TYPE "st_Io_Ph_DigitalOutputs"
VERSION : 0.1
   STRUCT
      Zone1_K7k5Ss_Close { ExternalAccessible := 'False'; ExternalVisible := 'False'; ExternalWritable := 'False'; S7_SetPoint := 'False'} : "st_Io_Ph_DigitalOutput";
      Zone1_K7k5Vfd_Close { ExternalAccessible := 'False'; ExternalVisible := 'False'; ExternalWritable := 'False'; S7_SetPoint := 'False'} : "st_Io_Ph_DigitalOutput";
      Zone1_K37Ss_Close { ExternalAccessible := 'False'; ExternalVisible := 'False'; ExternalWritable := 'False'; S7_SetPoint := 'False'} : "st_Io_Ph_DigitalOutput";
      Zone1_K37Vfd_Close { ExternalAccessible := 'False'; ExternalVisible := 'False'; ExternalWritable := 'False'; S7_SetPoint := 'False'} : "st_Io_Ph_DigitalOutput";
      Zone1_K110Ss_Close { ExternalAccessible := 'False'; ExternalVisible := 'False'; ExternalWritable := 'False'; S7_SetPoint := 'False'} : "st_Io_Ph_DigitalOutput";
      Zone1_K110Vfd_Close { ExternalAccessible := 'False'; ExternalVisible := 'False'; ExternalWritable := 'False'; S7_SetPoint := 'False'} : "st_Io_Ph_DigitalOutput";
      Zone1_Q560Ss_Open { ExternalAccessible := 'False'; ExternalVisible := 'False'; ExternalWritable := 'False'; S7_SetPoint := 'False'} : "st_Io_Ph_DigitalOutput";
      Zone1_Q560Ss_Close { ExternalAccessible := 'False'; ExternalVisible := 'False'; ExternalWritable := 'False'; S7_SetPoint := 'False'} : "st_Io_Ph_DigitalOutput";
      Zone1_Q560Ss_ChargeSpring { ExternalAccessible := 'False'; ExternalVisible := 'False'; ExternalWritable := 'False'; S7_SetPoint := 'False'} : "st_Io_Ph_DigitalOutput";
      Zone1_Q630Vfd_Open { ExternalAccessible := 'False'; ExternalVisible := 'False'; ExternalWritable := 'False'; S7_SetPoint := 'False'} : "st_Io_Ph_DigitalOutput";
      Zone1_Q630Vfd_Close { ExternalAccessible := 'False'; ExternalVisible := 'False'; ExternalWritable := 'False'; S7_SetPoint := 'False'} : "st_Io_Ph_DigitalOutput";
      Zone1_Q630Vfd_ChargeSpring { ExternalAccessible := 'False'; ExternalVisible := 'False'; ExternalWritable := 'False'; S7_SetPoint := 'False'} : "st_Io_Ph_DigitalOutput";
      Zone1_LampGreen { ExternalAccessible := 'False'; ExternalVisible := 'False'; ExternalWritable := 'False'; S7_SetPoint := 'False'} : "st_Io_Ph_DigitalOutput";
      Zone1_LampYellow { ExternalAccessible := 'False'; ExternalVisible := 'False'; ExternalWritable := 'False'; S7_SetPoint := 'False'} : "st_Io_Ph_DigitalOutput";
      Zone1_LampRed { ExternalAccessible := 'False'; ExternalVisible := 'False'; ExternalWritable := 'False'; S7_SetPoint := 'False'} : "st_Io_Ph_DigitalOutput";
      Zone1_LampStart { ExternalAccessible := 'False'; ExternalVisible := 'False'; ExternalWritable := 'False'; S7_SetPoint := 'False'} : "st_Io_Ph_DigitalOutput";
      Zone1_LampStop { ExternalAccessible := 'False'; ExternalVisible := 'False'; ExternalWritable := 'False'; S7_SetPoint := 'False'} : "st_Io_Ph_DigitalOutput";
      Zone1_LampTakeSample { ExternalAccessible := 'False'; ExternalVisible := 'False'; ExternalWritable := 'False'; S7_SetPoint := 'False'} : "st_Io_Ph_DigitalOutput";
      Zone1_LampEStop { ExternalAccessible := 'False'; ExternalVisible := 'False'; ExternalWritable := 'False'; S7_SetPoint := 'False'} : "st_Io_Ph_DigitalOutput";
      Zone1_LampPanelEStop { ExternalAccessible := 'False'; ExternalVisible := 'False'; ExternalWritable := 'False'; S7_SetPoint := 'False'} : "st_Io_Ph_DigitalOutput";
      Zone2_K7k5Ss_Close { ExternalAccessible := 'False'; ExternalVisible := 'False'; ExternalWritable := 'False'; S7_SetPoint := 'False'} : "st_Io_Ph_DigitalOutput";
      Zone2_K7k5Vfd_Close { ExternalAccessible := 'False'; ExternalVisible := 'False'; ExternalWritable := 'False'; S7_SetPoint := 'False'} : "st_Io_Ph_DigitalOutput";
      Zone2_K37Ss_Close { ExternalAccessible := 'False'; ExternalVisible := 'False'; ExternalWritable := 'False'; S7_SetPoint := 'False'} : "st_Io_Ph_DigitalOutput";
      Zone2_K37Vfd_Close { ExternalAccessible := 'False'; ExternalVisible := 'False'; ExternalWritable := 'False'; S7_SetPoint := 'False'} : "st_Io_Ph_DigitalOutput";
      Zone2_K110Ss_Close { ExternalAccessible := 'False'; ExternalVisible := 'False'; ExternalWritable := 'False'; S7_SetPoint := 'False'} : "st_Io_Ph_DigitalOutput";
      Zone2_K110Vfd_Close { ExternalAccessible := 'False'; ExternalVisible := 'False'; ExternalWritable := 'False'; S7_SetPoint := 'False'} : "st_Io_Ph_DigitalOutput";
      Zone2_Q560Ss_Open { ExternalAccessible := 'False'; ExternalVisible := 'False'; ExternalWritable := 'False'; S7_SetPoint := 'False'} : "st_Io_Ph_DigitalOutput";
      Zone2_Q560Ss_Close { ExternalAccessible := 'False'; ExternalVisible := 'False'; ExternalWritable := 'False'; S7_SetPoint := 'False'} : "st_Io_Ph_DigitalOutput";
      Zone2_Q560Ss_ChargeSpring { ExternalAccessible := 'False'; ExternalVisible := 'False'; ExternalWritable := 'False'; S7_SetPoint := 'False'} : "st_Io_Ph_DigitalOutput";
      Zone2_Q630Vfd_Open { ExternalAccessible := 'False'; ExternalVisible := 'False'; ExternalWritable := 'False'; S7_SetPoint := 'False'} : "st_Io_Ph_DigitalOutput";
      Zone2_Q630Vfd_Close { ExternalAccessible := 'False'; ExternalVisible := 'False'; ExternalWritable := 'False'; S7_SetPoint := 'False'} : "st_Io_Ph_DigitalOutput";
      Zone2_Q630Vfd_ChargeSpring { ExternalAccessible := 'False'; ExternalVisible := 'False'; ExternalWritable := 'False'; S7_SetPoint := 'False'} : "st_Io_Ph_DigitalOutput";
      Zone2_LampGreen { ExternalAccessible := 'False'; ExternalVisible := 'False'; ExternalWritable := 'False'; S7_SetPoint := 'False'} : "st_Io_Ph_DigitalOutput";
      Zone2_LampYellow { ExternalAccessible := 'False'; ExternalVisible := 'False'; ExternalWritable := 'False'; S7_SetPoint := 'False'} : "st_Io_Ph_DigitalOutput";
      Zone2_LampRed { ExternalAccessible := 'False'; ExternalVisible := 'False'; ExternalWritable := 'False'; S7_SetPoint := 'False'} : "st_Io_Ph_DigitalOutput";
      Zone2_LampStart { ExternalAccessible := 'False'; ExternalVisible := 'False'; ExternalWritable := 'False'; S7_SetPoint := 'False'} : "st_Io_Ph_DigitalOutput";
      Zone2_LampStop { ExternalAccessible := 'False'; ExternalVisible := 'False'; ExternalWritable := 'False'; S7_SetPoint := 'False'} : "st_Io_Ph_DigitalOutput";
      Zone2_LampTakeSample { ExternalAccessible := 'False'; ExternalVisible := 'False'; ExternalWritable := 'False'; S7_SetPoint := 'False'} : "st_Io_Ph_DigitalOutput";
      Zone2_LampEStop { ExternalAccessible := 'False'; ExternalVisible := 'False'; ExternalWritable := 'False'; S7_SetPoint := 'False'} : "st_Io_Ph_DigitalOutput";
      Zone2_LampPanelEStop { ExternalAccessible := 'False'; ExternalVisible := 'False'; ExternalWritable := 'False'; S7_SetPoint := 'False'} : "st_Io_Ph_DigitalOutput";
      Zone3_K7k5Ss_Close { ExternalAccessible := 'False'; ExternalVisible := 'False'; ExternalWritable := 'False'; S7_SetPoint := 'False'} : "st_Io_Ph_DigitalOutput";
      Zone3_K7k5Vfd_Close { ExternalAccessible := 'False'; ExternalVisible := 'False'; ExternalWritable := 'False'; S7_SetPoint := 'False'} : "st_Io_Ph_DigitalOutput";
      Zone3_K37Ss_Close { ExternalAccessible := 'False'; ExternalVisible := 'False'; ExternalWritable := 'False'; S7_SetPoint := 'False'} : "st_Io_Ph_DigitalOutput";
      Zone3_K37Vfd_Close { ExternalAccessible := 'False'; ExternalVisible := 'False'; ExternalWritable := 'False'; S7_SetPoint := 'False'} : "st_Io_Ph_DigitalOutput";
      Zone3_K110Ss_Close { ExternalAccessible := 'False'; ExternalVisible := 'False'; ExternalWritable := 'False'; S7_SetPoint := 'False'} : "st_Io_Ph_DigitalOutput";
      Zone3_K110Vfd_Close { ExternalAccessible := 'False'; ExternalVisible := 'False'; ExternalWritable := 'False'; S7_SetPoint := 'False'} : "st_Io_Ph_DigitalOutput";
      Zone3_Q560Ss_Open { ExternalAccessible := 'False'; ExternalVisible := 'False'; ExternalWritable := 'False'; S7_SetPoint := 'False'} : "st_Io_Ph_DigitalOutput";
      Zone3_Q560Ss_Close { ExternalAccessible := 'False'; ExternalVisible := 'False'; ExternalWritable := 'False'; S7_SetPoint := 'False'} : "st_Io_Ph_DigitalOutput";
      Zone3_Q560Ss_ChargeSpring { ExternalAccessible := 'False'; ExternalVisible := 'False'; ExternalWritable := 'False'; S7_SetPoint := 'False'} : "st_Io_Ph_DigitalOutput";
      Zone3_Q630Vfd_Open { ExternalAccessible := 'False'; ExternalVisible := 'False'; ExternalWritable := 'False'; S7_SetPoint := 'False'} : "st_Io_Ph_DigitalOutput";
      Zone3_Q630Vfd_Close { ExternalAccessible := 'False'; ExternalVisible := 'False'; ExternalWritable := 'False'; S7_SetPoint := 'False'} : "st_Io_Ph_DigitalOutput";
      Zone3_Q630Vfd_ChargeSpring { ExternalAccessible := 'False'; ExternalVisible := 'False'; ExternalWritable := 'False'; S7_SetPoint := 'False'} : "st_Io_Ph_DigitalOutput";
      Zone3_LampGreen { ExternalAccessible := 'False'; ExternalVisible := 'False'; ExternalWritable := 'False'; S7_SetPoint := 'False'} : "st_Io_Ph_DigitalOutput";
      Zone3_LampYellow { ExternalAccessible := 'False'; ExternalVisible := 'False'; ExternalWritable := 'False'; S7_SetPoint := 'False'} : "st_Io_Ph_DigitalOutput";
      Zone3_LampRed { ExternalAccessible := 'False'; ExternalVisible := 'False'; ExternalWritable := 'False'; S7_SetPoint := 'False'} : "st_Io_Ph_DigitalOutput";
      Zone3_LampStart { ExternalAccessible := 'False'; ExternalVisible := 'False'; ExternalWritable := 'False'; S7_SetPoint := 'False'} : "st_Io_Ph_DigitalOutput";
      Zone3_LampStop { ExternalAccessible := 'False'; ExternalVisible := 'False'; ExternalWritable := 'False'; S7_SetPoint := 'False'} : "st_Io_Ph_DigitalOutput";
      Zone3_LampTakeSample { ExternalAccessible := 'False'; ExternalVisible := 'False'; ExternalWritable := 'False'; S7_SetPoint := 'False'} : "st_Io_Ph_DigitalOutput";
      Zone3_LampEStop { ExternalAccessible := 'False'; ExternalVisible := 'False'; ExternalWritable := 'False'; S7_SetPoint := 'False'} : "st_Io_Ph_DigitalOutput";
      Zone3_LampPanelEStop { ExternalAccessible := 'False'; ExternalVisible := 'False'; ExternalWritable := 'False'; S7_SetPoint := 'False'} : "st_Io_Ph_DigitalOutput";
      Drive_7k5Ss_Run { ExternalAccessible := 'False'; ExternalVisible := 'False'; ExternalWritable := 'False'; S7_SetPoint := 'False'} : "st_Io_Ph_DigitalOutput";
      Drive_7k5Vfd_Run { ExternalAccessible := 'False'; ExternalVisible := 'False'; ExternalWritable := 'False'; S7_SetPoint := 'False'} : "st_Io_Ph_DigitalOutput";
      Drive_37Ss_Run { ExternalAccessible := 'False'; ExternalVisible := 'False'; ExternalWritable := 'False'; S7_SetPoint := 'False'} : "st_Io_Ph_DigitalOutput";
      Drive_37Vfd_Run { ExternalAccessible := 'False'; ExternalVisible := 'False'; ExternalWritable := 'False'; S7_SetPoint := 'False'} : "st_Io_Ph_DigitalOutput";
      Drive_110Ss_Run { ExternalAccessible := 'False'; ExternalVisible := 'False'; ExternalWritable := 'False'; S7_SetPoint := 'False'} : "st_Io_Ph_DigitalOutput";
      Drive_110Vfd_Run { ExternalAccessible := 'False'; ExternalVisible := 'False'; ExternalWritable := 'False'; S7_SetPoint := 'False'} : "st_Io_Ph_DigitalOutput";
      Drive_560Ss_Run { ExternalAccessible := 'False'; ExternalVisible := 'False'; ExternalWritable := 'False'; S7_SetPoint := 'False'} : "st_Io_Ph_DigitalOutput";
      Drive_630Vfd_Run { ExternalAccessible := 'False'; ExternalVisible := 'False'; ExternalWritable := 'False'; S7_SetPoint := 'False'} : "st_Io_Ph_DigitalOutput";
   END_STRUCT;

END_TYPE

